{attribute 'qualified_only'}

VAR_GLOBAL RETAIN
	GeneralSwitchConfig : stSwitchConfig :=(ShortClickMaxTime := T#300MS,
									ShortClickDelayTime := T#400MS,
									LongClickMaxTime := T#1000MS);
									
END_VAR

(* stored: Version 1.1.0.1
   GVL gvlSwitches: Id {e6e0d0e9-0431-466b-ba2e-1acdfc72ee46} *)
